// TIA Portal project "REMPLISSAGE DES CUVES D'EAU" (V16)

(* hardware
DEVICE "Station S7-1200_1"  S7-1200 Station
   slot 0: "Châssis_0"  S7-1200 Rack  Rack  V1.0
   slot 1: "PLC_1"  CPU 1214C AC/DC/Rly  6ES7 214-1BG40-0XB0  V4.4
*)

// ===== PLC "PLC_1"  CPU 1214C AC/DC/Rly =====

VAR_GLOBAL   // PLC tag table "Table de variables standard"
   "BP_S1" AT %I0.0 : Bool;
   "BP_STOP" AT %I0.1 : Bool;
   "NHH1" AT %M0.2 : Bool;
   "MARCHE_SYS" AT %M0.3 : Bool;
END_VAR

ORGANIZATION_BLOCK "Main"   // OB1, LAD, ProgramCycle
TITLE = "Main Program Sweep (Cycle)" / PROGRAMME DE REMPLISSAGE DES CUVES
{ S7_Optimized_Access := 'TRUE' }
VERSION : 0.1
   VAR_INPUT
      Initial_Call : Bool;   // Initial call of this OB
      Remanence : Bool;   // =True, if remanent data are available
   END_VAR
BEGIN

REGION Network 1: MARCHE/ARRET
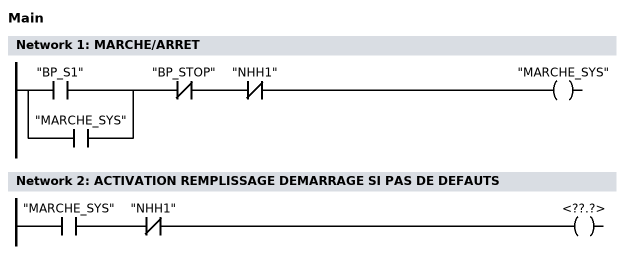
   RUNG wire#powerrail
      Contact( "BP_S1" )
      wire#w1
      I_Contact( "BP_STOP" )
      I_Contact( "NHH1" )
      Coil( "MARCHE_SYS" )
   END_RUNG
   RUNG wire#powerrail
      Contact( "MARCHE_SYS" )
   END_RUNG wire#w1
   // the same network as SCL:
   "MARCHE_SYS" := ("BP_S1" OR "MARCHE_SYS") AND NOT "BP_STOP" AND NOT "NHH1";
END_REGION

REGION Network 2: ACTIVATION REMPLISSAGE DEMARRAGE SI PAS DE DEFAUTS
   RUNG wire#powerrail
      Contact( "MARCHE_SYS" )
      I_Contact( "NHH1" )
      Coil(  )
   END_RUNG
   // the same network as SCL:
   <??.?> := "MARCHE_SYS" AND NOT "NHH1";
END_REGION
END_ORGANIZATION_BLOCK